Fanuc KAREL source: KT00425.KL

PROGRAM KT00425
%NOLOCKGROUP
VAR
  P1: XYZWPR
  P2: XYZWPREXT
  OUT: BOOLEAN
BEGIN
  P1.X = 1.0
    P2.Y = 2.0
  OUT = P1 > P2
END KT00425
